FUNCTION_BLOCK FB_Element// EXTENDS FB_SFC_Cycle IMPLEMENTS ITF_FB_SFC_Cycle
VAR_INPUT
	eElementID			: E_Element_List;

END_VAR
VAR_OUTPUT
	event_StateUpdate	: INT; // for HMI
END_VAR



VAR
	eType				: E_Element_Type;
	eProdType			: E_Product_Type;
	eState_Long			: E_Element_State_Long;
	eState_Short		: E_Element_State_Short;
	eState_Long_last	: E_Element_State_Long;
	eState_Long_Expiered: E_Element_State_Long;





	i: INT;
	sState_Time			: STRING;
	sTimeToExpiration	: STRING;
	tTimeToExpiration	: TIME;
	tStateTime			: TIME;

	
	sElementID			: STRING;
	eInterConnect		: E_InterConnection;
	memoDissolving_active		: BOOL;
	bStateUpdate_Limited		: BOOL;

	stCIP_Request		: ST_CIP_Request;
	stCIP_RequestActive	: ST_CIP_Request;

	bTakePosInCIPBuffer_Partial		: BOOL;
	bTakePosInCIPBuffer_Full		: BOOL;
	bTakePosInCIPBuffer_Detergent	: BOOL;
	bError: BOOL;	
	
	eProdStatus			: E_Prod_Status;
	eFilling_State		: E_Filling_State;
	
	fbEvent_echo: FB_Event_echo;

END_VAR

VAR PERSISTENT
	tsStateChange				: TimeStruct;
	tsCIP						: TimeStruct;
	tsWater						: TimeStruct;
	tsProduction				: TimeStruct;
	tsProductionLine			: TimeStruct;
	tsProductionLineStby		: TimeStruct;
	
	
	tExpirationTime				: TIME:=T#48H;
	ExDuration_Product			: TIME:=T#48H; 	//Expiration from loaded ricipe
	ExDuration_Water			: TIME:=T#48H; 	//Expiration from loaded ricipe
	
	eExTime						: E_ExTime;


END_VAR


VAR_IN_OUT
	stOperation		: ST_OperationButtons;	
END_VAR

i:=i+1;
//m_Set_SFCFlags_Reference();
//SUPER^();
fbEvent_echo(echo=>event_StateUpdate);
act_StateMachine();
act_StateChange_WatchGog();

sElementID:=TO_STRING(eElementID);

CASE eType OF 
	E_Element_Type.eTank:;
				act_Tank();
	E_Element_Type.eTriBlender:;
				act_TriBlender();
	E_Element_Type.eLine:;
				act_Line();

END_CASE

CASE eElementID OF
	E_Element_List.eTank_1:;
				eType:=E_Element_Type.eTank;
				eProdType:=E_Product_Type.Marinada;
				stCIP_Request.eClient:=E_CIP_Usage.eTank_1;
	E_Element_List.eTank_2:;
				eType:=E_Element_Type.eTank;
				eProdType:=E_Product_Type.Marinada;
				stCIP_Request.eClient:=E_CIP_Usage.eTank_2;
	E_Element_List.eTank_3:;
				eType:=E_Element_Type.eTank;
				eProdType:=E_Product_Type.Color;
				stCIP_Request.eClient:=E_CIP_Usage.eTank_3;
	E_Element_List.eTank_4:;
				eType:=E_Element_Type.eTank;
				eProdType:=E_Product_Type.Color;
				stCIP_Request.eClient:=E_CIP_Usage.eTank_4;
	E_Element_List.eTriBlender_Marinada:;
				eType:=E_Element_Type.eTriBlender;
				eProdType:=E_Product_Type.Marinada;		
				stCIP_Request.eClient:=E_CIP_Usage.eTriBlender_Marinada;
	E_Element_List.eTriBlender_Color:;
				eType:=E_Element_Type.eTriBlender;
				eProdType:=E_Product_Type.Color;
				stCIP_Request.eClient:=E_CIP_Usage.eTriBlender_Color;
	E_Element_List.eLine_Marinada:;
				eType:=E_Element_Type.eLine;
				eProdType:=E_Product_Type.Marinada;
				stCIP_Request.eClient:=E_CIP_Usage.eLine_Marinada;
	E_Element_List.eLine_Color:;
				eType:=E_Element_Type.eLine;
				eProdType:=E_Product_Type.Color;
				stCIP_Request.eClient:=E_CIP_Usage.eLine_Color;
END_CASE


IF bTakePosInCIPBuffer_Partial THEN;
	stCIP_Request.eType:=E_CIP_Type.R_Water;
	fbCIP.m_TakePosInCIPBuffer(stCIP_Request:=stCIP_Request);
	bTakePosInCIPBuffer_Partial:=FALSE;
END_IF

IF bTakePosInCIPBuffer_Detergent THEN;
	stCIP_Request.eType:=E_CIP_Type.Detergent;
	fbCIP.m_TakePosInCIPBuffer(stCIP_Request:=stCIP_Request);
	bTakePosInCIPBuffer_Detergent:=FALSE;
END_IF

IF bTakePosInCIPBuffer_Full THEN;
	stCIP_Request.eType:=E_CIP_Type.Full;
	fbCIP.m_TakePosInCIPBuffer(stCIP_Request:=stCIP_Request);
	bTakePosInCIPBuffer_Full:=FALSE;
END_IF

stCIP_RequestActive.eType:=E_CIP_Type.NotSelected;
FOR i:=0 TO 9 DO
	IF arCIP_RequestBufer[i].eClient=stCIP_Request.eClient
	AND arCIP_RequestBufer[i].eType>stCIP_RequestActive.eType THEN;
		stCIP_RequestActive.eType:=arCIP_RequestBufer[i].eType;
	END_IF
END_FOR

m_TimeToExpiration();

ACTION act_Line:

END_ACTION

ACTION act_StateChange_WatchGog:
IF eState_Long<>eState_Long_last THEN;
	IF eState_Long=E_Element_State_Long.eExpired THEN;
		eState_Long_Expiered:=eState_Long_last;
	ELSE;
		eState_Long_Expiered:=E_Element_State_Long.eOff;
	END_IF

	IF eState_Long=E_Element_State_Long.eWaterReady THEN;
		IF  eState_Long_last=E_Element_State_Long.eCIP_5_Done THEN;
			//tsWater:=stSystemTime;
			m_Set_TimeToExpirationMode(eExTime_set:=E_ExTime.eWater);
		ELSE;
			// do nothing here...
		END_IF
		
	ELSIF eState_Long>=E_Element_State_Long.eReady THEN;
		IF eState_Long=E_Element_State_Long.eReady
		AND NOT memoDissolving_active THEN; // state updated manualy
			m_Set_Dissolveng_active_memo();
		ELSE; // state update during dissolving status
			// do nothing here...
		END_IF
	ELSE;
		//tsCIP:=stSystemTime;
		m_Set_TimeToExpirationMode(eExTime_set:=E_ExTime.eCIP);
		
	END_IF
	
	eState_Long_last:=eState_Long;
	
	fbEvent_echo.event(); // for HMI
END_IF

tStateTime:=TO_TIME(SYSTEMTIME_TO_DT(stSystemTime)-SYSTEMTIME_TO_DT(tsStateChange));

sState_Time:=prg_RealClock.m_DeltaTime(stStartTime:=tsStateChange);
sTimeToExpiration:=prg_RealClock.mTime_to_String_HMI(tInputTime:=tTimeToExpiration, iSecondDisplay:=TRUE);

sState_Time:= CONCAT(sState_Time, '(');
sState_Time:= CONCAT(sState_Time, sTimeToExpiration);
sState_Time:= CONCAT(sState_Time, ')');

CASE eExTime OF 
	E_ExTime.eCIP:sState_Time:= CONCAT(sState_Time, '/C');
	E_ExTime.eLine:sState_Time:= CONCAT(sState_Time, '/L');
	E_ExTime.eLineStby:sState_Time:= CONCAT(sState_Time, '/LS');
	E_ExTime.eProduct:sState_Time:= CONCAT(sState_Time, '/P');
	E_ExTime.eWater:sState_Time:= CONCAT(sState_Time, '/W');
	
END_CASE
END_ACTION

ACTION act_StateMachine:
CASE eState_Long OF
	E_Element_State_Long.eOff,
	E_Element_State_Long.eStandby,
	E_Element_State_Long.eNotClean,
	E_Element_State_Long.eCIP_1_Rinzed,
	E_Element_State_Long.eCIP_2_Deterged,
	E_Element_State_Long.eCIP_3_Deterged_Clean,	
	E_Element_State_Long.eCIP_4_Sanitized:;
				eState_Short:=E_Element_State_Short.eNotClean;
					ExpirationTime:=ExDuration_Default;
	E_Element_State_Long.eCIP_5_Done:;
				eState_Short:=E_Element_State_Short.eClean;
					memoDissolving_active:=FALSE;
	E_Element_State_Long.eWaterReady:;	
				IF memoDissolving_active THEN;
					eState_Short:=E_Element_State_Short.eProduct;
				ELSE;
					eState_Short:=E_Element_State_Short.eClean;
				END_IF
	E_Element_State_Long.eReady,
	E_Element_State_Long.eProduction,
	E_Element_State_Long.eEmpty:;	
				eState_Short:=E_Element_State_Short.eProduct;
	E_Element_State_Long.eExpired:;
				//
	
END_CASE
END_ACTION

ACTION act_Tank:
;
END_ACTION

ACTION act_TriBlender:
(*
IF eInterConnect=E_InterConnection.ConnToCIP 
AND eElementID=E_Element_List.eTriBlender_Marinada
AND eTriBlenderPipe<>E_TriBlenderPipe.eMarinada
THEN;
	bError:=TRUE;
ELSE;
	bError:=FALSE;
END_IF
*)
END_ACTION

PROPERTY ExpirationMode : E_ExTime
GET
ExpirationMode:=eExTime;
END_GET
SET
eExTime:=ExpirationMode;
END_SET
END_PROPERTY

PROPERTY ExpirationTime : TIME
GET
ExpirationTime:=tExpirationTime;
END_GET
SET
tExpirationTime:=ExpirationTime;
END_SET
END_PROPERTY

PROPERTY Interconnect : E_InterConnection
GET
Interconnect:=m_Get_InterConnection();
END_GET
SET
END_SET
END_PROPERTY

METHOD m_Disconnect : BOOL
VAR_INPUT
END_VAR
eInterConnect:=E_InterConnection.NotConnected;
CASE eType OF
	E_Element_Type.eTank:;					
			//
	E_Element_Type.eTriBlender,
	E_Element_Type.eLine:;
			//tsProductionLineStby:=stSystemTime;
			m_Set_TimeToExpirationMode(eExTime_set:=E_ExTime.eLineStby);
END_CASE
END_METHOD

METHOD m_Get_CIP_Avilable : BOOL
VAR_INPUT
END_VAR
IF TRUE 
AND (eInterConnect=E_InterConnection.NotConnected OR eInterConnect=E_InterConnection.ConnToCIP)
AND TRUE
THEN;
	m_Get_CIP_Avilable:=TRUE;
ELSE;
	m_Get_CIP_Avilable:=FALSE;
END_IF
END_METHOD

METHOD m_Get_InterConnection : E_InterConnection
VAR_INPUT
END_VAR

m_Get_InterConnection:=eInterConnect;
END_METHOD

METHOD m_Get_Oper_Pause_Puls : BOOL
VAR_INPUT
END_VAR
m_Get_Oper_Pause_Puls:=stOperation.b_rt_Pause;
END_METHOD

METHOD m_Get_Oper_Pause_State : BOOL
VAR_INPUT
END_VAR
IF stOperation.b_rt_Pause THEN;
	m_Get_Oper_Pause_State:=TRUE;
ELSE;
	m_Get_Oper_Pause_State:=FALSE;
END_IF
END_METHOD

METHOD m_Get_Oper_Play_Puls : BOOL
VAR_INPUT
END_VAR
m_Get_Oper_Play_Puls:=stOperation.b_rt_Play;
END_METHOD

METHOD m_Get_Oper_Play_State : BOOL
VAR_INPUT
END_VAR
IF stOperation.iActOperation=E_OperationButtons.ePlayAll THEN;
	m_Get_Oper_Play_State:=TRUE;
ELSE;
	m_Get_Oper_Play_State:=FALSE;
END_IF
END_METHOD

METHOD m_Get_State : E_Element_State_Long
VAR_INPUT
END_VAR
m_Get_State:=eState_Long;
END_METHOD

METHOD m_Get_State_Short : E_Element_State_Short
VAR_INPUT
END_VAR
m_Get_State_Short:=eState_Short;
END_METHOD

METHOD m_Get_TimeToExpirationMode : TIME
VAR_INPUT
	eExTime_check		: E_ExTime;
END_VAR

VAR
	tsStateChange_local				: TimeStruct;
	tModeTime		: TIME;
	tModeDuration	: TIME;

END_VAR
CASE eExTime_check OF
	E_ExTime.eCIP:;
			tsStateChange_local:=tsCIP;
			tModeDuration:=ExDuration_Default;
	E_ExTime.eWater:;
			tsStateChange_local:=tsWater;
			tModeDuration:=ExDuration_Water;
	E_ExTime.eProduct:;
			tsStateChange_local:=tsProduction;	
			tModeDuration:=ExDuration_Product;
	E_ExTime.eLine :;
			tsStateChange_local:=tsProductionLine;
			tModeDuration:=ExDuration_Default_Line;
	E_ExTime.eLineStby:;
			tsStateChange_local:=tsProductionLineStby;
			tModeDuration:=ExDuration_Default_LineStandby;
END_CASE
tModeTime:=TO_TIME(SYSTEMTIME_TO_DT(stSystemTime)-SYSTEMTIME_TO_DT(tsStateChange_local));
m_Get_TimeToExpirationMode:=tModeDuration-tModeTime;
END_METHOD

METHOD m_Get_Type : E_Element_Type
VAR_INPUT
END_VAR
m_Get_Type:=eType;
END_METHOD

METHOD m_InterConnect : BOOL
VAR_INPUT
	value: E_InterConnection;
END_VAR
IF eInterConnect=E_InterConnection.NotConnected 
OR eInterConnect=value
THEN;
	eInterConnect:=value;
	m_InterConnect:=TRUE;
ELSE;
	m_InterConnect:=FALSE;
END_IF
END_METHOD

METHOD m_InterConnected_State : BOOL
VAR_INPUT
	eState_Long_Set			: E_Element_State_Long;
END_VAR

IF (eState_Long_Set>eState_Long 
OR eState_Long_Set=E_Element_State_Long.eNotClean)
AND eState_Long_Set<=E_Element_State_Long.eProduction
THEN;
	eState_Long:=eState_Long_Set;
END_IF
END_METHOD

METHOD m_Set_Dissolveng_active_memo : BOOL
VAR_INPUT
END_VAR
IF NOT memoDissolving_active THEN;
	
	
	IF eInterConnect=E_InterConnection.ConnToTank THEN;
		//tsProductionLine:=stSystemTime;
		m_Set_TimeToExpirationMode(eExTime_set:=E_ExTime.eLine);
	ELSE; //element is production tank
		//tsProduction:=stSystemTime;
		m_Set_TimeToExpirationMode(eExTime_set:=E_ExTime.eProduct);
	END_IF
	
END_IF
memoDissolving_active:=TRUE;
fbEvent_echo.event();
END_METHOD

METHOD m_Set_ExpirationDuration : BOOL
VAR_INPUT
	eExTime_set		: E_ExTime;
	setTime			: TIME;

END_VAR
CASE eExTime_set OF
	E_ExTime.eCIP:;
			
	E_ExTime.eWater:;
			ExDuration_Water:=setTime;
			m_Set_ExpirationDuration:=TRUE;
	E_ExTime.eProduct:;
			ExDuration_Product:=setTime;	
			m_Set_ExpirationDuration:=TRUE;
	E_ExTime.eLine :;
			
	E_ExTime.eLineStby:;
			
END_CASE
END_METHOD

METHOD m_Set_Oper_Pause
VAR_INPUT
END_VAR
IF stOperation.iActOperation<>E_OperationButtons.ePauseAll THEN;
	stOperation.bSetPause:=TRUE;
END_IF
END_METHOD

METHOD m_Set_Oper_Play
VAR_INPUT
END_VAR
IF stOperation.iActOperation<>E_OperationButtons.ePlayAll THEN;
	stOperation.bSetPlay:=TRUE;
END_IF
END_METHOD

METHOD m_Set_SFCFlags_Reference : BOOL
//Set reference to SFC flags

refSFC.SFCInit REF= SFCInit;
refSFC.SFCReset REF= SFCReset;
refSFC.SFCError REF= SFCError;
refSFC.SFCEnableLimit REF= SFCEnableLimit;
refSFC.SFCErrorStep REF= SFCErrorStep;
refSFC.SFCErrorPOU REF= SFCErrorPOU;
refSFC.SFCQuitError REF= SFCQuitError;
refSFC.SFCPause REF= SFCPause;
refSFC.SFCTrans REF= SFCTrans;
refSFC.SFCCurrentStep REF= SFCCurrentStep;
refSFC.SFCTip REF= SFCTip;
refSFC.SFCTipMode REF= SFCTipMode;

// Cycle handle for SFC
m_SFC_Handle();
END_METHOD

METHOD m_Set_State : BOOL
VAR_INPUT
	eState_Long_Set			: E_Element_State_Long;
END_VAR
(*
IF eState_Long_Set>eState_Long 
OR eState_Long_Set=E_Element_State_Long.eNotClean
THEN;
	eState_Long:=eState_Long_Set;
END_IF
*)
eState_Long:=eState_Long_Set;
END_METHOD

METHOD m_Set_TimeToExpirationMode : TIME
VAR_INPUT
	eExTime_set		: E_ExTime;
END_VAR

VAR
	tsSet				: TimeStruct;
	tsStateChange_local				: TimeStruct;
	tModeTime		: TIME;
	tModeDuration	: TIME;

END_VAR
tsSet:=stSystemTime;
CASE eExTime_set OF
	E_ExTime.eCIP:;
			tsStateChange_local:=tsCIP:=tsSet;
			tModeDuration:=ExDuration_Default;
	E_ExTime.eWater:;
			tsStateChange_local:=tsWater:=tsSet;
			tModeDuration:=ExDuration_Water;
	E_ExTime.eProduct:;
			tsStateChange_local:=tsProduction:=tsSet;	
			tModeDuration:=ExDuration_Product;
	E_ExTime.eLine :;
			tsStateChange_local:=tsProductionLine:=tsSet;
			tModeDuration:=ExDuration_Default_Line;
	E_ExTime.eLineStby:;
			tsStateChange_local:=tsProductionLineStby:=tsSet;
			tModeDuration:=ExDuration_Default_LineStandby;
END_CASE
tModeTime:=TO_TIME(SYSTEMTIME_TO_DT(stSystemTime)-SYSTEMTIME_TO_DT(tsStateChange_local));
m_Set_TimeToExpirationMode:=tModeDuration-tModeTime;

CASE eExTime OF
	E_ExTime.eCIP:;
			tsStateChange:=tsCIP;
	E_ExTime.eWater:;
			tsStateChange:=tsWater;
	E_ExTime.eProduct:;
			tsStateChange:=tsProduction;			
	E_ExTime.eLine :;
			tsStateChange:=tsProductionLine;
	E_ExTime.eLineStby:;
			tsStateChange:=tsProductionLineStby;
END_CASE
END_METHOD

METHOD m_StateUpdate_Limit : BOOL
VAR_INPUT
	value: BOOL;
END_VAR
IF value THEN;
	bStateUpdate_Limited:=TRUE;
ELSE;
	bStateUpdate_Limited:=FALSE;
END_IF
END_METHOD

METHOD m_TimeExpiered : BOOL
VAR_INPUT
END_VAR
CASE eType OF
	E_Element_Type.eTank:;			
	E_Element_Type.eTriBlender:;
	E_Element_Type.eLine:;
	
END_CASE
	
// Rolling Down option
CASE eInterConnect OF
	E_InterConnection.NotConnected:;
				m_TimeExpiredState_RollDown();
	E_InterConnection.ConnToCIP:;
				//do nothing
	E_InterConnection.ConnToLine,
	E_InterConnection.ConnToTriBlender:;
				// Type Tank
				m_TimeExpiredState_RollDown();
	E_InterConnection.ConnToTank:;
				//do nothing
	
END_CASE
END_METHOD

METHOD m_TimeExpiredState_RollDown : BOOL
VAR_INPUT
END_VAR
CASE eState_Long OF
	E_Element_State_Long.eCIP_1_Rinzed:;
				//
	E_Element_State_Long.eCIP_2_Deterged,
	E_Element_State_Long.eCIP_3_Deterged_Clean,
	E_Element_State_Long.eCIP_4_Sanitized,
	E_Element_State_Long.eCIP_5_Done:;	
				State:=E_Element_State_Long.eCIP_1_Rinzed;
	E_Element_State_Long.eWaterReady,
	E_Element_State_Long.eReady,
	E_Element_State_Long.eProduction,
	E_Element_State_Long.eEmpty:;	
			IF eType=E_Element_Type.eTank THEN;
				//State:=E_Element_State_Long.eExpired;
				CASE eElementID OF 
					E_Element_List.eTank_1:;
						IF fbTank1.bReady THEN;
							State:=E_Element_State_Long.eExpired;
						END_IF
						
					E_Element_List.eTank_2:;
						IF fbTank2.bReady THEN;
							State:=E_Element_State_Long.eExpired;
						END_IF
						
					E_Element_List.eTank_3:;
						IF fbTank3.bReady THEN;
							State:=E_Element_State_Long.eExpired;
						END_IF
						
					E_Element_List.eTank_4:;
						IF fbTank4.bReady THEN;
							State:=E_Element_State_Long.eExpired;
						END_IF
												
				END_CASE
				
			ELSE;
				State:=E_Element_State_Long.eNotClean;
			END_IF
			
		E_Element_State_Long.eExpired:;
				IF eType=E_Element_Type.eLine OR eType=E_Element_Type.eTriBlender THEN;
					State:=E_Element_State_Long.eNotClean;
				END_IF
END_CASE
END_METHOD

METHOD m_TimeToExpiration : BOOL
VAR_INPUT
END_VAR
IF tExpirationTime>tStateTime THEN;
	tTimeToExpiration:=tExpirationTime-tStateTime;
ELSE;
	tTimeToExpiration:=T#0S;
	IF TRUE 
	AND eFilling_State=E_Filling_State.eFilling_InProcess
	AND eType=E_Element_Type.eTank
	AND eInterConnect <> E_InterConnection.NotConnected
	AND TRUE
	THEN;
		//Production filling in process 
	ELSE;
		m_TimeExpiered();
	END_IF
	
END_IF

IF State=E_Element_State_Long.eExpired THEN;
	m_TimeExpiered();	
END_IF

IF State=E_Element_State_Long.eStandby 
OR State=E_Element_State_Long.eNotClean
THEN;
	tTimeToExpiration:=T#0S;
END_IF


CASE eType OF
	E_Element_Type.eTank:;		
			CASE eState_Short OF
				E_Element_State_Short.eNotClean:;
						ExpirationTime:=ExDuration_Default;
						eExTime:=E_ExTime.eCIP;
				E_Element_State_Short.eClean:;
						IF eState_Long=E_Element_State_Long.eWaterReady 
						OR (eState_Long=E_Element_State_Long.eExpired
							AND eState_Long_Expiered=E_Element_State_Long.eWaterReady)
						THEN;
							ExpirationTime:=ExDuration_Water;
							eExTime:=E_ExTime.eWater;
						ELSE;
							ExpirationTime:=ExDuration_Default;
							eExTime:=E_ExTime.eCIP;
						END_IF
				E_Element_State_Short.eProduct:;
						ExpirationTime:=ExDuration_Product;
						eExTime:=E_ExTime.eProduct;
			END_CASE			
			
	E_Element_Type.eTriBlender,
	E_Element_Type.eLine:;
			CASE eInterConnect OF
				E_InterConnection.NotConnected:;
					CASE eState_Short OF
						E_Element_State_Short.eNotClean,
						E_Element_State_Short.eClean:;
								ExpirationTime:=ExDuration_Default;
								eExTime:=E_ExTime.eCIP;
	
						E_Element_State_Short.eProduct:;
								IF m_Get_TimeToExpirationMode(eExTime_check:=E_ExTime.eLine)<ExDuration_Default_LineStandby THEN; // line remain time less then 2 hours
									ExpirationTime:=ExDuration_Default_Line;
									eExTime:=E_ExTime.eLine;
								ELSE;
									ExpirationTime:=ExDuration_Default_LineStandby;
									eExTime:=E_ExTime.eLineStby;
								END_IF								
					END_CASE
			
				E_InterConnection.ConnToCIP:;
						ExpirationTime:=ExDuration_Default;
						eExTime:=E_ExTime.eCIP;
						
				E_InterConnection.ConnToTank:;
					CASE eState_Short OF
						E_Element_State_Short.eNotClean,
						E_Element_State_Short.eClean:;
								ExpirationTime:=ExDuration_Default;
								eExTime:=E_ExTime.eCIP;
	
						E_Element_State_Short.eProduct:;		
								ExpirationTime:=ExDuration_Default_Line;
								eExTime:=E_ExTime.eLine;				
					END_CASE
	
						
			ELSE;
		END_CASE
END_CASE


CASE eExTime OF
	E_ExTime.eCIP:;
			tsStateChange:=tsCIP;
	E_ExTime.eWater:;
			tsStateChange:=tsWater;
	E_ExTime.eProduct:;
			tsStateChange:=tsProduction;			
	E_ExTime.eLine :;
			tsStateChange:=tsProductionLine;
	E_ExTime.eLineStby:;
			tsStateChange:=tsProductionLineStby;
END_CASE

CASE eInterConnect OF
	E_InterConnection.NotConnected:;
	E_InterConnection.ConnToCIP:;
	E_InterConnection.ConnToTank:;
	E_InterConnection.ConnToLine:;
	E_InterConnection.ConnToTriBlender:;
END_CASE
END_METHOD

PROPERTY pFilling_State : E_Filling_State
GET
pFilling_State:=eFilling_State;
END_GET
SET
eFilling_State:=pFilling_State;
END_SET
END_PROPERTY

PROPERTY ProdStatus : E_Prod_Status
GET
ProdStatus:=eProdStatus;
END_GET
SET
eProdStatus:=ProdStatus;
END_SET
END_PROPERTY

PROPERTY State : E_Element_State_Long
GET
State:=eState_Long;
END_GET
SET
eState_Long:=State;
END_SET
END_PROPERTY

PROPERTY StateTime : TIMESTRUCT
GET
StateTime:=tsStateChange;
END_GET
SET

CASE eState_Long OF 
	E_Element_State_Long.eOff..			
	E_Element_State_Long.eCIP_5_Done:;
				tsStateChange:=StateTime;
				
				
	//E_Element_State_Long.eOff:;
	//E_Element_State_Long.eOff:;
	//E_Element_State_Long.eOff:;
	
END_CASE
END_SET
END_PROPERTY

END_FUNCTION_BLOCK

(* stored: Version 1.1.0.1, ProductVersion 3.1.4024.15
   POU FB_Element: Id {700358c5-37aa-4b9c-88fa-65bcc8fcf7eb}, SpecialFunc None
   Folder Manage: Id {c1bad6aa-d321-46fa-921e-00f6b446e0b8}
   Folder Property: Id {aa60355e-95fb-4f4a-adf9-1e47dcacbd8b}
   Action act_Line: Id {7224f2cd-9678-4b86-88f6-72fd19bfe71e}
   Action act_StateChange_WatchGog: Id {4dafd2ba-8022-4674-a1d5-a6952dfd70bd}
   Action act_StateMachine: Id {f33c6159-2800-4ae4-981a-4a8c5e4774dd}
   Action act_Tank: Id {2dddeb0d-68bf-4477-8840-0824af0883b1}
   Action act_TriBlender: Id {26031c10-f211-4816-a500-dc05d95c74de}
   Property ExpirationMode: Id {e272ce08-3353-4f37-8b69-bb279f090906}
   Get Get: Id {6f2c38fe-4df9-472f-aa93-91c22dd94c80}
   Set Set: Id {8ef68865-931e-45f9-90dd-d20b3c5e284e}
   Property ExpirationTime: Id {2df3d745-ae6c-40b9-bacc-a56f4fe0173c}
   Get Get: Id {1b57346c-44cd-46d9-8e51-18e302aa4b85}
   Set Set: Id {1a5c7ea4-8b69-46ee-b373-941be47f8b05}
   Property Interconnect: Id {59358565-33fe-4169-84cb-6ec04b788a77}
   Get Get: Id {e7f086bb-f260-4468-a17a-f433c6eed49e}
   Set Set: Id {f2915f05-4763-4ad6-b220-04929851b8fb}
   Method m_Disconnect: Id {20e4c919-f24b-4fbd-ae5c-73c93cc7bd42}
   Method m_Get_CIP_Avilable: Id {85fd739d-7b69-4185-bc50-898d5ccfd7e4}
   Method m_Get_InterConnection: Id {b128ae88-6959-4ba2-8ec6-647a3af8a375}
   Method m_Get_Oper_Pause_Puls: Id {d59793fd-b3de-47f1-8e51-0b1c0e5d5b3f}
   Method m_Get_Oper_Pause_State: Id {a2cc3607-da54-4c2f-b052-7ea6fd6c809c}
   Method m_Get_Oper_Play_Puls: Id {57c42df4-a06a-4bc2-8394-7fb8c54c97b4}
   Method m_Get_Oper_Play_State: Id {1d8040a3-b691-4499-92e8-a729d8801f54}
   Method m_Get_State: Id {54c18fb6-79a0-4507-a1ae-52b2474932d3}
   Method m_Get_State_Short: Id {a4895e89-8af5-4844-8a6f-98d623177713}
   Method m_Get_TimeToExpirationMode: Id {d304daf3-a250-4e31-b078-0f17be3d063d}
   Method m_Get_Type: Id {e3e31f5e-e6b1-403c-bb2b-b2d06d0264ea}
   Method m_InterConnect: Id {72ff53e2-bb5f-4090-a2e6-ef10be06eb5a}
   Method m_InterConnected_State: Id {c4bb22d1-79f1-477b-b979-1591791ba3b1}
   Method m_Set_Dissolveng_active_memo: Id {55ab6cb4-4a2f-4aab-971f-9547041e4c7f}
   Method m_Set_ExpirationDuration: Id {d852322c-ba1c-43fa-ac6b-bcfdfd4889f5}
   Method m_Set_Oper_Pause: Id {31bfa777-0c86-4838-93b6-ec28e092b686}
   Method m_Set_Oper_Play: Id {6a6aba07-12dd-441c-945b-5a5009b81ef4}
   Method m_Set_SFCFlags_Reference: Id {173e8058-adb0-4138-b5d3-8a3b87ec3293}
   Method m_Set_State: Id {5873be97-3110-49a4-84ea-a94cd608159b}
   Method m_Set_TimeToExpirationMode: Id {b4162e1c-9425-4a9c-aebb-53e10584e3d9}
   Method m_StateUpdate_Limit: Id {fb1d1185-6118-48f5-8cfa-978fe0325d17}
   Method m_TimeExpiered: Id {0e06182a-e09e-4ec2-920d-88b3137754d2}
   Method m_TimeExpiredState_RollDown: Id {2f9443d7-fd06-45c2-8331-f1b6d4473c16}
   Method m_TimeToExpiration: Id {b592f2a7-8b80-4b25-9040-91bd7248992a}
   Property pFilling_State: Id {3fb22dff-576a-4883-be93-9c6c846c05ea}
   Get Get: Id {479b8e08-02fe-4667-920d-886fec9827b0}
   Set Set: Id {3f3e119f-2905-4e48-a771-ff3266f5ea5f}
   Property ProdStatus: Id {e4474016-ac40-43b2-890c-a624cfadb69e}
   Get Get: Id {d8c98c4f-e4a7-4d29-8f1c-e4501e77bc63}
   Set Set: Id {493fd571-f83e-4f1f-9bab-25e613c526d3}
   Property State: Id {b7a48a0b-d269-4423-aeca-a5757298ed3c}
   Get Get: Id {72cbb051-9d79-4c21-a7db-ea4f457a68c7}
   Set Set: Id {a5ff53c4-2a1a-43d5-8777-6503e1925952}
   Property StateTime: Id {93f72989-6112-490b-ac1e-9957a7069cbd}
   Get Get: Id {806b7699-7a09-4a45-b13d-b3d26a5a904b}
   Set Set: Id {79374df6-a9bd-428c-a0c7-b15c90bc1b1d} *)
